Staubli VAL3: logicIF.pgx

public program logicIF(num x_nResult1, num x_nResult2, num x_nResult3, bool x_bANDOR1, bool x_bANDOR2, bool& x_bFinalResult)
  local bool l_bFinalResult1
  local bool l_bFinalResult2
begin
  if x_nResult1==0 and x_nResult2==0 and x_nResult3==0
    x_bFinalResult=false
  elseIf x_nResult1==0 and x_nResult2==0 and x_nResult3!=0
    x_bFinalResult=(x_nResult3==1)
  elseIf x_nResult1==0 and x_nResult2!=0 and x_nResult3==0
    x_bFinalResult=(x_nResult2==1)
  elseIf x_nResult1!=0 and x_nResult2==0 and x_nResult3==0
    x_bFinalResult=(x_nResult1==1)
  elseIf x_nResult1!=0 and x_nResult2!=0 and x_nResult3==0
    if x_bANDOR1
      x_bFinalResult=(x_nResult1==1 or x_nResult2==1)
    else
      x_bFinalResult=(x_nResult1==1 and x_nResult2==1)
    endIf
  elseIf x_nResult1==0 and x_nResult2!=0 and x_nResult3!=0
    if x_bANDOR2
      x_bFinalResult=(x_nResult1==1 or x_nResult2==1)
    else
      x_bFinalResult=(x_nResult1==1 and x_nResult2==1)
    endIf
  elseIf x_nResult1!=0 and x_nResult2!=0 and x_nResult3!=0
    if x_bANDOR1 and x_bANDOR2
      x_bFinalResult=(x_nResult1==1 or x_nResult2==1 or x_nResult3==1)
    elseIf !x_bANDOR1 and !x_bANDOR2
      x_bFinalResult=(x_nResult1==1 and x_nResult2==1 and x_nResult3==1)
    elseIf !x_bANDOR1 and x_bANDOR2
      x_bFinalResult=(x_nResult1==1 and x_nResult2==1 or x_nResult3==1)
    elseIf x_bANDOR1 and !x_bANDOR2
      x_bFinalResult=((x_nResult1==1 or x_nResult2==1) and x_nResult3==1)
    endIf

  endIf
end
